FUNCTION_BLOCK SingleActingActuator (* Basic Function Block Type *)
  (* Standard: 61499-2 *)
  (* Version 0.0, 7/2/2026, Template *)
  PACKAGE Main;
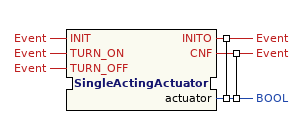
  EVENT_INPUT
    INIT; (* Initialization Request *)
    TURN_ON; (* Normal Execution Request *)
    TURN_OFF;
  END_EVENT
  EVENT_OUTPUT
    INITO WITH actuator; (* Initialization Confirm *)
    CNF WITH actuator; (* Execution Confirmation *)
  END_EVENT
  VAR_OUTPUT
    actuator : BOOL; (* Output event qualifier *)
  END_VAR
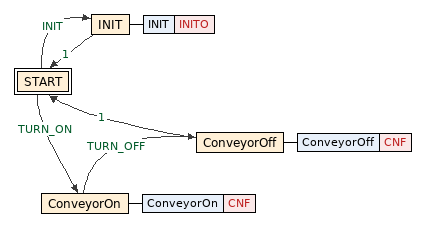
  EC_STATES
    START; (* Initial State *)
    INIT : INIT -> INITO; (* Initialization *)
    ConveyorOff : ConveyorOff -> CNF;
    ConveyorOn : ConveyorOn -> CNF;
  END_STATES
  EC_TRANSITIONS
    START TO INIT := INIT;
    INIT TO START := 1;
    START TO ConveyorOn := TURN_ON;
    ConveyorOff TO START := 1;
    ConveyorOn TO ConveyorOff := TURN_OFF;
  END_TRANSITIONS
  ALGORITHM INIT IN ST: (* Initialization algorithm *)
actuator := FALSE;
  END_ALGORITHM
  ALGORITHM REQ IN ST: (* Normally executed algorithm *)
;
  END_ALGORITHM
  ALGORITHM ConveyorOn IN ST:
actuator := TRUE;
  END_ALGORITHM
  ALGORITHM ConveyorOff IN ST:
actuator := FALSE;
  END_ALGORITHM
END_FUNCTION_BLOCK
